Staubli VAL3: clearActStack.pgx

public program clearActStack()
  local num l_n
begin
  for l_n=0 to size(_nPuleStartClk)-1
    _nPuleStartClk[l_n]=-1
  endFor
  _nActStackIndex=0
  for l_n=0 to size(actCmd)-1
    call removeActCmd(l_n)
  endFor
end
